(* IEC 61131-3 sources: trust-platform/examples/filling_line/src, 7 files *)

(* ---- Types.st ---- *)
TYPE
    E_Mode : (Stopped, Filling, Draining);
END_TYPE

(* ---- Interfaces.st ---- *)
INTERFACE IValve
    METHOD Open : BOOL
    END_METHOD

    METHOD Close : BOOL
    END_METHOD

    PROPERTY IsOpen : BOOL
        GET
        END_GET
    END_PROPERTY
END_INTERFACE

INTERFACE IPump
    METHOD Start : BOOL
    END_METHOD

    METHOD Stop : BOOL
    END_METHOD

    PROPERTY IsRunning : BOOL
        GET
        END_GET
    END_PROPERTY

    PROPERTY Speed : INT
        GET
        END_GET
        SET
        END_SET
    END_PROPERTY
END_INTERFACE

(* ---- LevelControllerFb.st ---- *)
FUNCTION_BLOCK LevelControllerFb2
VAR_INPUT
    LevelPct : REAL;
    StartCmd : BOOL;
    StopCmd : BOOL;
END_VAR
VAR_OUTPUT
    FillCmd : BOOL;
    DrainCmd : BOOL;
    Mode : E_Mode;
END_VAR
VAR
    target : REAL := 70.0;
    hysteresis : REAL := 5.0;
END_VAR

IF StopCmd THEN
    Mode := E_Mode#Stopped;
ELSIF StartCmd THEN
    IF LevelPct < target - hysteresis THEN
        Mode := E_Mode#Filling;
    ELSIF LevelPct > target + hysteresis THEN
        Mode := E_Mode#Draining;
    ELSE
        Mode := E_Mode#Stopped;
    END_IF;
END_IF;

FillCmd := Mode = E_Mode#Filling;
DrainCmd := Mode = E_Mode#Draining;
END_FUNCTION_BLOCK

(* ---- PumpFb.st ---- *)
FUNCTION_BLOCK PumpFb IMPLEMENTS IPump
VAR
    running : BOOL;
    speed_value : INT;
END_VAR

METHOD PUBLIC Start : BOOL
    running := TRUE;
    Start := running;
END_METHOD

METHOD PUBLIC Stop : BOOL
    running := FALSE;
    Stop := running;
END_METHOD

PUBLIC PROPERTY IsRunning : BOOL
    GET
        IsRunning := running;
    END_GET
    SET
    END_SET
END_PROPERTY

PUBLIC PROPERTY Speed : INT
    GET
        Speed := speed_value;
    END_GET
    SET
        speed_value := Speed;
    END_SET
END_PROPERTY
END_FUNCTION_BLOCK

(* ---- ValveFb.st ---- *)
FUNCTION_BLOCK ValveFb IMPLEMENTS IValve
VAR
    open_state : BOOL;
END_VAR

METHOD PUBLIC Open : BOOL
    open_state := TRUE;
    Open := open_state;
END_METHOD

METHOD PUBLIC Close : BOOL
    open_state := FALSE;
    Close := open_state;
END_METHOD

PUBLIC PROPERTY IsOpen : BOOL
    GET
        IsOpen := open_state;
    END_GET
END_PROPERTY
END_FUNCTION_BLOCK

(* ---- Configuration.st ---- *)
CONFIGURATION FillingLine
TASK Cycle (INTERVAL := T#50ms, PRIORITY := 1);
PROGRAM P1 WITH Cycle : MainProgram;
VAR_CONFIG
    P1.StartCmd AT %IX0.0 : BOOL;
    P1.StopCmd AT %IX0.1 : BOOL;
    P1.LevelRaw AT %IW0 : INT;
    P1.FillValveOut AT %QX0.0 : BOOL;
    P1.DrainValveOut AT %QX0.1 : BOOL;
    P1.PumpSpeedOut AT %QW0 : INT;
END_VAR
END_CONFIGURATION

(* ---- Main.st ---- *)
PROGRAM MainProgram
VAR
    StartCmd : BOOL;
    StopCmd : BOOL;
    LevelRaw : INT;
    FillValveOut : BOOL;
    DrainValveOut : BOOL;
    PumpSpeedOut : INT;

    LevelPct : REAL;
    Ctrl : LevelControllerFb2;
END_VAR

LevelPct := INT_TO_REAL(LevelRaw) * 0.1;

Ctrl(LevelPct := LevelPct, StartCmd := StartCmd, StopCmd := StopCmd);

IF Ctrl.FillCmd THEN
    FillValveOut := TRUE;
    DrainValveOut := FALSE;
    PumpSpeedOut := INT#800;
ELSIF Ctrl.DrainCmd THEN
    FillValveOut := FALSE;
    DrainValveOut := TRUE;
    PumpSpeedOut := INT#600;
ELSE
    FillValveOut := FALSE;
    DrainValveOut := FALSE;
    PumpSpeedOut := INT#0;
END_IF;
END_PROGRAM
